(* Logix 5000 project; controller MECO9497 vendor 1 type 14 code 106 rev 21.11; software revision 21.00 *)

TASK MainTask (continuous, watchdog 500 ms) : MainProgram
TASK PID_LOOP (periodic, rate 250 ms, priority 5, watchdog 500 ms) : PID_MAIN
TASK PID_SLOW (periodic, rate 1000 ms, priority 10, watchdog 500 ms) : PID_SLOW

MODULES
   Local : vendor 1 type 14 code 106 (Compact 0, rev 21.11)
       : 1769-IQ16 (Compact 1, rev 1.1, Input RPI 20 ms)
       : 1769-IF8 (Compact 3, rev 1.1, Output RPI 80 ms)
       : vendor 1 type 10 code 40 (Compact 5, rev 2.1, Output RPI 80 ms)
       : 1769-OW16 (Compact 2, rev 1.1, Output RPI 20 ms)
       : 1769-IF8 (Compact 4, rev 1.1, Output RPI 80 ms)
END_MODULES

VAR_GLOBAL   (* controller tags *)
   AAH_200 : BOOL := 1;
   AAH_200_ACK : BOOL;
   AAH_200_AUX : BOOL := 1;
   AAH_200_DELAY : TIMER := (PRE := 1000);
   AAH_200_DI : ALIAS FOR Local:1:I.Data.5;
   AAH_200_SP : REAL := 0.6;
   AAH_200_SP_H : BOOL;
   AAH_200_SP_N : BOOL;
   AAH_200_SP_O : REAL := 0.6;
   ACKNOWLEDGE : BOOL;
   ALARM_ACK_OIT : BOOL;
   ALARM_HORN_DO : ALIAS FOR Local:2:O.Data.10;
   ALARM_RESET_OIT : BOOL;
   ALARM_SCREEN_DISPLAY_BIT : BOOL;
   ALARM_SCREEN_LATCH_BIT : BOOL;
   ALERT_ALARM_SU_DELAY : TIMER := (PRE := 300000);
   ALERT_ALARM_SU_DELAY_H : BOOL;
   ALERT_ALARM_SU_DELAY_N : BOOL;
   ALERT_ALARM_SU_DELAY_O : DINT := 300;
   AT_200_AI : ALIAS FOR Local:4:I.Ch0Data;
   AT_200_EU : REAL;
   AUDIBLE_SUMMARY : BOOL;
   COMP_AMP_ALRM_DELAY_TMR : TIMER := (PRE := 20000);
   COMP_BUMP_OIT : BOOL;
   COMP_BUMP_SU_DELAY : TIMER := (PRE := 20);
   COMPRESSOR_FAULT_DELAY : TIMER := (PRE := 3000);
   COMPRESSOR_MOTOR_FLT_STARTUP_DELAY : TIMER := (PRE := 6000);
   COMPRESSOR_MOTOR_START_DELAY : TIMER := (PRE := 5000);
   COMPRESSOR_MOTOR_START_DO : ALIAS FOR Local:2:O.Data.0;
   COMPRESSOR_START_CMD : BOOL;
   CR_4 : ALIAS FOR Local:2:O.Data.9;
   CR_6 : ALIAS FOR Local:2:O.Data.2;
   CURRENT_SCREEN : DINT := 7;
   D_V_ALERT_ALARM : BOOL;
   D_V_CRITICAL_ALARM : BOOL;
   D_V_OP_SWITCH_AUTO : BOOL := 1;
   D_V_OP_SWITCH_MAN : BOOL;
   D_V_OP_SWITCH_OFF : BOOL;
   D_V_REMOTE_START : BOOL;
   D_V_REMOTE_START_MAP : BOOL;
   D_V_UNIT_RUNNIING : BOOL;
   DELTA_V_FP : REAL[30] := ([2] := 0.006103888, [4] := 0.25801086, [5] := 100.0, [6] := 60.074467, [8] := 39.310135, [9] := 1.5030825, [11] := 40.0, [12] := 102.87493, [13] := 102.08753); {produced}
   DELTA_V_READ : INT[10] := ([0] := 2, [2] := 1344, [3] := 16383, [5] := 1); {produced}
   DELTA_V_WRITE : INT[10] := ([0] := 1); {produced}
   DIST_COND_ALRM_STARTUP_TIME_H : BOOL;
   DIST_COND_ALRM_STARTUP_TIME_N : BOOL;
   DIST_COND_ALRM_STARTUP_TIME_O : REAL := 300.0;
   DIST_COND_ALRM_STARTUP_TMR : TIMER := (PRE := 300000);
   DIST_MOTOR_BUMP_OIT : BOOL;
   DIST_PUMP_START_SP : REAL := 75.0;
   DIST_PUMP_START_SP_H : BOOL;
   DIST_PUMP_START_SP_N : BOOL;
   DIST_PUMP_START_SP_OIT : REAL := 80.0;
   DIST_PUMP_STOP_SP : REAL := 10.0;
   DIST_PUMP_STOP_SP_H : BOOL;
   DIST_PUMP_STOP_SP_N : BOOL;
   DIST_PUMP_STOP_SP_OIT : DINT := 20;
   DIST_TO_STORAGE_TIME_SP_H : BOOL;
   DIST_TO_STORAGE_TIME_SP_N : BOOL;
   DIST_TO_STORAGE_TIME_SP_OIT : DINT;
   DISTILATE_TO_STORAGE : BOOL;
   DISTILLATE_MOTOR_FAULT_DELAY : TIMER := (PRE := 3000);
   DISTILLATE_MOTOR_START_DO : ALIAS FOR Local:2:O.Data.1;
   DISTILLATE_PUMP_NORM_START : BOOL;
   DISTILLATE_PUMP_START_CMD : BOOL;
   DISTILLATE_PUMP_STDBY_START : BOOL;
   DSTLT_BOX_DRAIN_HOT_STANDBY : TIMER := (PRE := 600000, ACC := 600000, EN := 1, DN := 1);
   DSTLT_BOX_DRAIN_HOT_STANDBY_CLOSE : TIMER := (PRE := 1800000, ACC := 431720, EN := 1, TT := 1);
   DSTLT_BOX_DRAIN_NORM_DELAY : TIMER := (PRE := 5000);
   DSTLT_BOX_DRAIN_STANDBY : BOOL;
   DSTLT_BOX_DRAIN_STBY_DELAY_TIMER : TIMER := (PRE := 10000);
   DSTLT_PUMP_START_DELAY : TIMER := (PRE := 5000);
   DSTLT_PUMP_STBY_STOP_SP : REAL;
   DSTLT_PUMP_STBY_STRT_SP : REAL;
   DSTLT_STORAGE : BOOL;
   DSTLT_STORAGE_DELAY_TIMER : TIMER := (PRE := 60000);
   DSTLT_STORAGE_DELTA_V : BOOL;
   DSTLT_STORAGE_ENABLE_MAP : BOOL := 1;
   DSTLT_STORAGE_ENABLE_OIT : BOOL := 1;
   DSTLT_TEMP_ALRM_SU_DELAY : TIMER := (PRE := 300000);
   DSTLT_TEMP_ALRM_SU_DELAY_H : BOOL;
   DSTLT_TEMP_ALRM_SU_DELAY_N : BOOL;
   DSTLT_TEMP_ALRM_SU_DELAY_O : REAL := 300.0;
   DSTLT_TEMP_CNTRL_DELAY_TIMER : TIMER := (PRE := 90000);
   E_Stop : ALIAS FOR Local:1:I.Data.0;
   E_Stop_ACK : BOOL;
   E_Stop_AUX : BOOL := 1;
   E_Stop_DI_MAP : BOOL;
   ENGINEER : BOOL;
   EVAP_PRESS_CV_LIMIT : BOOL;
   EVAP_PRESS_CV_PERMISSIVE : REAL := 10.0;
   EVAP_PRESS_RAMP_ONE_SHOT : BOOL;
   EVAP_PRESS_RAMP_TIMER : TIMER := (PRE := 60000);
   EVAP_PRESSURE_CV_PERM : BOOL := 1;
   EVAP_PRESSURE_PERM : BOOL := 1;
   EVAP_PRESSURE_PERM_TIME_H : BOOL;
   EVAP_PRESSURE_PERM_TIME_N : BOOL;
   EVAP_PRESSURE_PERM_TIME_O : REAL := 180.0;
   EVAP_PRESSURE_PERM_TIMER : TIMER := (PRE := 180000, ACC := 180000, EN := 1, DN := 1);
   EVAP_RAMP_COMPLETE : BOOL;
   EVAP_RAMP_ENABLE_DELAY_TIMER : TIMER := (PRE := 180000);
   EXCESS_DIST_TIME_SP_H : BOOL;
   EXCESS_DIST_TIME_SP_N : BOOL;
   EXCESS_DIST_TIME_SP_OIT : REAL := 10.0;
   EXCESS_DIST_TO_DRAIN_ACK : BOOL;
   EXCESS_DIST_TO_DRAIN_AUX : BOOL := 1;
   EXCESS_DSTLT_DELAY_TIMER : TIMER := (PRE := 1000);
   EXCESS_DSTLT_DRAIN : BOOL := 1;
   EXCESS_DSTLT_DRAIN_TIMER : TIMER := (PRE := 600000);
   EXCESS_DSTLT_REMAIN : DINT := 10;
   FC_300_AM_OIT : BOOL;
   FC_300_OS_OFF : BOOL := 1;
   FC_300_OS_ON : BOOL;
   FC_300_SP : DINT := 58;
   FC_300_SP_H : BOOL;
   FC_300_SP_N : BOOL;
   FC_300_SP_O : DINT := 58;
   FC_300_SP_OUT : DINT;
   FEED_LVL_CV_LIMIT : BOOL := 1;
   FEED_LVL_CV_LIMIT_SHUTDOWN : BOOL := 1;
   FEED_LVL_CV_LIMIT_SHUTDOWN_DELAY : TIMER := (PRE := 30000);
   FEED_LVL_CV_LIMIT_SHUTDOWN_LATCH : BOOL;
   FEED_LVL_ONE_SHOT : BOOL;
   FEED_TEM_SD_LATCH : BOOL;
   FEED_TEM_SD_TIMER : TIMER := (PRE := 30000);
   FEED_TEMP_SD_ONS : BOOL := 1;
   FEED_TEMP_STEP_DELAY : TIMER := (PRE := 10000);
   FT_200_AI : ALIAS FOR Local:3:I.Ch2Data;
   FT_200_EU : REAL;
   HEARTBEAT : BOOL := 1;
   HEARTBEAT_AUX : BOOL;
   HEARTBEAT_OUT : BOOL := 1;
   HEARTBEAT_RESET_OIT : BOOL;
   HOT_STANDBY : BOOL := 1;
   HOURMETER_DO : ALIAS FOR Local:2:O.Data.4;
   IAL_100 : BOOL;
   IAL_100_ACK : BOOL;
   IAL_100_AUX : BOOL := 1;
   IAL_100_CTR : COUNTER := (PRE := 3);
   IAL_100_DELAY : TIMER := (PRE := 5000);
   IAL_100_SP : REAL := 30.0;
   IAL_100_SP_H : BOOL;
   IAL_100_SP_N : BOOL;
   IAL_100_SP_OIT : REAL := 30.0;
   INITIAL_SCAN_BIT : BOOL;
   INITIAL_SCAN_SYS_RESET : BOOL;
   INITIAL_SCAN_SYS_RESET_TMR : TIMER := (PRE := 30000);
   INITIAL_START_STEAM_LIMIT_TMR : TIMER := (PRE := 300000, ACC := 300000, EN := 1, DN := 1);
   IY_100_AI : ALIAS FOR Local:4:I.Ch2Data;
   IY_100_EU : REAL;
   LAAH_100 : BOOL := 1;
   LAAH_100_ACK : BOOL;
   LAAH_100_ALERT_H : BOOL;
   LAAH_100_ALERT_N : BOOL;
   LAAH_100_ALERT_O : DINT := 80;
   LAAH_100_AUX : BOOL := 1;
   LAAH_100_DELAY : TIMER := (PRE := 5000);
   LAAH_100_SP : DINT := 80;
   LAAL_100 : BOOL := 1;
   LAAL_100_ACK : BOOL;
   LAAL_100_ALERT_H : BOOL;
   LAAL_100_ALERT_N : BOOL;
   LAAL_100_ALERT_O : DINT := 20;
   LAAL_100_AUX : BOOL := 1;
   LAAL_100_DELAY : TIMER := (PRE := 1000);
   LAAL_100_SP : DINT := 20;
   LAH_100 : BOOL := 1;
   LAH_100_ACK : BOOL;
   LAH_100_AUX : BOOL := 1;
   LAH_100_DELAY : TIMER := (PRE := 5000);
   LAH_100_SP : REAL := 80.0;
   LAH_100_SP_H : BOOL;
   LAH_100_SP_N : BOOL;
   LAH_100_SP_OIT : REAL := 80.0;
   LAL_100 : BOOL := 1;
   LAL_100_ACK : BOOL;
   LAL_100_AUX : BOOL := 1;
   LAL_100_DELAY : TIMER := (PRE := 1000);
   LAL_100_SP : REAL := 20.0;
   LAL_100_SP_H : BOOL;
   LAL_100_SP_N : BOOL;
   LAL_100_SP_OIT : REAL := 20.0;
   LATCH : BOOL := 1;
   LB_OIL_LOW_PRESS_ALRM_DELAY : TIMER := (PRE := 20000);
   LCV_100_AO : ALIAS FOR Local:5:O.Ch2Data;
   LCV_100_IND : DINT;
   LCV_100_INTERLOCK : BOOL := 1;
   LCV_200_AO : ALIAS FOR Local:5:O.Ch3Data;
   LCV_200_IND : DINT := 3;
   LIC_100 : PID := (CTL := -2139061120, EN := 1, PE := 1, INI := 1, DVNA := 1, PVHA := 1, SP := 9829.8, KP := 4.0, KI := 1.6, KD := 0.01, BIAS := -181.60863, MAXS := 16383.0, SO := 0.25801086, MAXO := 40.0, UPD := 0.25, PV := 9845.0, ERR := -15.200195, OUT := 0.25801086, MAXI := 16383.0, MAXCV := 16383.0, MAXTIE := 16383.0, DATA[0] := 182.52715, DATA[1] := -961.19507, DATA[2] := 9845.0, DATA[3] := -15.200195, DATA[4] := 9829.8, DATA[5] := 0.006103888, DATA[6] := 1.0, DATA[7] := 6.3999996, DATA[8] := 4.0, DATA[9] := 1.6, DATA[10] := 0.01, DATA[11] := 4.0, DATA[12] := 0.041666668, DATA[13] := 2.3999999, DATA[15] := 163.83, DATA[16] := 0.006103888);
   LIC_1000_CV1 : REAL := 20.0;
   LIC_100_A_M_OIT : BOOL;
   LIC_100_CV2 : REAL := 40.0;
   LIC_100_CV_H : BOOL;
   LIC_100_CV_N : BOOL;
   LIC_100_CV_OIT : REAL := 0.25801086;
   LIC_100_FINAL_SP : REAL := 9829.8;
   LIC_100_FINAL_SP_EU : REAL := 60.0;
   LIC_100_GAIN_H : BOOL;
   LIC_100_GAIN_N : BOOL;
   LIC_100_GAIN_OIT : REAL := 4.0;
   LIC_100_RATE_H : BOOL;
   LIC_100_RATE_N : BOOL;
   LIC_100_RATE_OIT : REAL := 0.01;
   LIC_100_RESET_H : BOOL;
   LIC_100_RESET_N : BOOL;
   LIC_100_RESET_OIT : REAL := 1.6;
   LIC_100_SP_CONV : REAL := 163.83;
   LIC_100_SP_EU : REAL := 60.0;
   LIC_100_SP_H : BOOL;
   LIC_100_SP_N : BOOL;
   LIC_100_SP_OIT : REAL := 60.0;
   LIC_100_STBY_SP : REAL := 9829.8;
   LIC_100_STBY_SP_EU : REAL := 60.0;
   LIC_100_STBY_SP_H : BOOL;
   LIC_100_STBY_SP_N : BOOL;
   LIC_100_STBY_SP_OIT : REAL := 60.0;
   LIC_200 : PID := (CTL := -2038397696, EN := 1, SWM := 1, CA := 1, PE := 1, INI := 1, DVNA := 1, PVLA := 1, SP := 9829.8, KP := 2.0, KI := 1.1, KD := 0.01, BIAS := 151.65573, MAXS := 16383.0, SO := 100.0, MAXO := 100.0, UPD := 0.25, PV := -98.0, ERR := -9927.8, OUT := 100.0, MAXI := 16383.0, MAXCV := 16383.0, MAXTIE := 16383.0, DATA[0] := 69.54062, DATA[1] := -9.570896, DATA[2] := -98.0, DATA[3] := -9927.8, DATA[4] := 9829.8, DATA[5] := 0.006103888, DATA[6] := 1.0, DATA[7] := 5.2, DATA[8] := 2.0, DATA[9] := 1.1, DATA[10] := 0.01, DATA[11] := 2.0, DATA[12] := 0.030303031, DATA[13] := 1.1999999, DATA[15] := 163.83, DATA[16] := 0.006103888);
   LIC_200_A_M_OIT : BOOL;
   LIC_200_CV_H : BOOL;
   LIC_200_CV_N : BOOL;
   LIC_200_CV_OIT : REAL := 100.0;
   LIC_200_GAIN_H : BOOL;
   LIC_200_GAIN_N : BOOL;
   LIC_200_GAIN_OIT : REAL := 2.0;
   LIC_200_RATE_H : BOOL;
   LIC_200_RATE_N : BOOL;
   LIC_200_RATE_OIT : REAL := 0.01;
   LIC_200_RESET_H : BOOL;
   LIC_200_RESET_N : BOOL;
   LIC_200_RESET_OIT : REAL := 1.1;
   LIC_200_SP_CONV : REAL := 163.83;
   LIC_200_SP_EU : REAL := 60.0;
   LIC_200_SP_H : BOOL;
   LIC_200_SP_N : BOOL;
   LIC_200_SP_OIT : REAL := 60.0;
   LT_100_AI : ALIAS FOR Local:3:I.Ch3Data;
   LT_100_EU : REAL := 60.092777;
   LT_100_EU_SPAN : REAL := 100.0;
   LT_100_EU_ZERO : REAL;
   LT_200_AI : ALIAS FOR Local:3:I.Ch4Data;
   LT_200_EU : REAL;
   LT_200_EU_SPAN : REAL := 100.0;
   LT_200_EU_ZERO : REAL;
   LUBE_OIL_PUMP_FAULT_DELAY : TIMER := (PRE := 3000);
   LUBE_OIL_PUMP_START_CMD : BOOL;
   LUBE_OIL_SHUTDWN_TIMER : TIMER := (PRE := 45000, ACC := 45000, EN := 1, DN := 1);
   M1_DI : ALIAS FOR Local:1:I.Data.1;
   M1_DI_MAP : BOOL;
   M1_FAULT_ACK : BOOL;
   M1_FAULT_AUX : BOOL := 1;
   M2_DI : ALIAS FOR Local:1:I.Data.2;
   M2_DI_MAP : BOOL;
   M2_FAULT_ACK : BOOL;
   M2_FAULT_AUX : BOOL := 1;
   M4_DI : ALIAS FOR Local:1:I.Data.4;
   M4_DI_MAP : BOOL;
   M4_FAULT_ACK : BOOL;
   M4_FAULT_AUX : BOOL := 1;
   MAINTENANCE : BOOL;
   MCB : BOOL;
   MSG_AAH_200 : BOOL;
   MSG_E_STOP : BOOL;
   MSG_EXCESS_DIST_TO_DRAIN : BOOL;
   MSG_IAL_100 : BOOL;
   MSG_LAH_100 : BOOL;
   MSG_LAL_100 : BOOL;
   MSG_M1_FLT : BOOL;
   MSG_M2_FLT : BOOL;
   MSG_M4_FLT : BOOL;
   MSG_PAH_103 : BOOL;
   MSG_PAL_103 : BOOL;
   MSG_PAL_700 : BOOL;
   MSG_TAH_700 : BOOL;
   MSG_TAL_200 : BOOL;
   MSS_ALERT : BOOL;
   MSS_AUTO_SHUTDOWN_LATCH : BOOL;
   MSS_SHUTDOWN : BOOL := 1;
   MSS_START_PERM : BOOL := 1;
   no : BOOL;
   OFF : BOOL;
   OIL_MOTOR_START_DO : ALIAS FOR Local:2:O.Data.11;
   OIT_SCREEN_CONTROL : DINT;
   OIT_SECURITY_LEVEL : DINT;
   OP_SWTCH_AUTO_DI : ALIAS FOR Local:1:I.Data.14;
   OP_SWTCH_AUTO_DI_MAP : BOOL := 1;
   OP_SWTCH_MANUAL_DI : ALIAS FOR Local:1:I.Data.13;
   OP_SWTCH_MANUAL_DI_MAP : BOOL;
   OPERATOR : BOOL;
   PAAH_103 : BOOL := 1;
   PAAH_103_ACK : BOOL;
   PAAH_103_ALERT_H : BOOL;
   PAAH_103_ALERT_N : BOOL;
   PAAH_103_ALERT_O : REAL := 3.0;
   PAAH_103_AUX : BOOL := 1;
   PAAH_103_DELAY : TIMER := (PRE := 1000);
   PAAH_103_SP : REAL := 3.0;
   PAAL_103 : BOOL := 1;
   PAAL_103_ACK : BOOL;
   PAAL_103_ALERT_H : BOOL;
   PAAL_103_ALERT_N : BOOL;
   PAAL_103_ALERT_O : REAL := 0.25;
   PAAL_103_AUX : BOOL := 1;
   PAAL_103_DELAY : TIMER := (PRE := 1000);
   PAAL_103_SP : REAL := 0.25;
   PAH_103 : BOOL := 1;
   PAH_103_ACK : BOOL;
   PAH_103_AUX : BOOL := 1;
   PAH_103_DELAY : TIMER := (PRE := 1000);
   PAH_103_SP : REAL := 3.0;
   PAH_103_SP_H : BOOL;
   PAH_103_SP_N : BOOL;
   PAH_103_SP_OIT : REAL := 3.0;
   PAL_103 : BOOL := 1;
   PAL_103_ACK : BOOL;
   PAL_103_AUX : BOOL := 1;
   PAL_103_DELAY : TIMER := (PRE := 1000);
   PAL_103_SP : REAL := 0.19;
   PAL_103_SP_H : BOOL;
   PAL_103_SP_N : BOOL;
   PAL_103_SP_OIT : REAL := 0.19;
   PAL_700 : BOOL;
   PAL_700_ACK : BOOL;
   PAL_700_ALRM_DELAY : TIMER := (PRE := 1000);
   PAL_700_AUX : BOOL := 1;
   PCV_103_AO : ALIAS FOR Local:5:O.Ch0Data;
   PCV_103_IND : DINT := 3;
   PCV_103_INTERLOCK : BOOL := 1;
   PERM_TIME_REMAINING : REAL;
   PIC_103 : PID := (CTL := -2139061120, EN := 1, PE := 1, INI := 1, DVNA := 1, PVHA := 1, SP := 4914.9004, KP := 3.5, KI := 1.0, KD := 0.01, BIAS := -117.88922, MAXS := 16383.0, SO := 39.310135, MAXO := 100.0, UPD := 0.25, PV := 4920.0, ERR := -5.0996094, OUT := 39.310135, MAXI := 16383.0, MAXCV := 16383.0, MAXTIE := 16383.0, DATA[0] := 157.11327, DATA[1] := -480.6931, DATA[2] := 4920.0, DATA[3] := -5.0996094, DATA[4] := 4914.9004, DATA[5] := 0.006103888, DATA[6] := 1.0, DATA[7] := 6.1, DATA[8] := 3.5, DATA[9] := 1.0, DATA[10] := 0.01, DATA[11] := 3.5, DATA[12] := 0.058333334, DATA[13] := 2.1, DATA[15] := 163.83, DATA[16] := 0.006103888);
   PIC_103_A_M_OIT : BOOL;
   PIC_103_CV_H : BOOL;
   PIC_103_CV_N : BOOL;
   PIC_103_CV_OIT : REAL := 38.848907;
   PIC_103_FINAL_SP : REAL := 1.0;
   PIC_103_GAIN_H : BOOL;
   PIC_103_GAIN_N : BOOL;
   PIC_103_GAIN_OIT : REAL := 3.5;
   PIC_103_RATE_H : BOOL;
   PIC_103_RATE_N : BOOL;
   PIC_103_RATE_OIT : REAL := 0.01;
   PIC_103_RESET_H : BOOL;
   PIC_103_RESET_N : BOOL;
   PIC_103_RESET_OIT : REAL := 1.0;
   PIC_103_SP_CONV : REAL := 3276.6;
   PIC_103_SP_EU : REAL := 1.5000001;
   PIC_103_SP_H : BOOL;
   PIC_103_SP_N : BOOL;
   PIC_103_SP_OIT : REAL := 1.0;
   PIC_103_STBY_SP : REAL := 4914.9004;
   PIC_103_STBY_SP_EU : REAL := 1.5000001;
   PIC_103_STBY_SP_H : BOOL;
   PIC_103_STBY_SP_N : BOOL;
   PIC_103_STBY_SP_OIT : REAL := 1.5;
   PSL_700_DI : ALIAS FOR Local:1:I.Data.7;
   PT_103_AI : ALIAS FOR Local:3:I.Ch0Data;
   PT_103_EU : REAL := 1.5015565;
   PT_103_EU_SPAN : REAL := 5.0;
   PT_103_EU_ZERO : REAL;
   PT_103_HIGH : REAL := 2.1;
   RESET : BOOL;
   RESET_CONDUCTIVITY_HIGH_OIT : BOOL;
   RESET_DIST_LOW_TEMP_OIT : BOOL;
   SECURITY_ENABLED : BOOL;
   SUPERVISOR : BOOL;
   SV_200 : ALIAS FOR Local:2:O.Data.5;
   SV_200_201_DO : ALIAS FOR Local:2:O.Data.6;
   SV_200_201_IND : BOOL;
   SV_200_CTL : BOOL;
   SV_200_IND : BOOL;
   SV_202_DO : ALIAS FOR Local:2:O.Data.5;
   SV_300_DO : ALIAS FOR Local:2:O.Data.3;
   SV_300_IND : BOOL;
   SV_500_DO : ALIAS FOR Local:2:O.Data.8;
   SV_500_IND : BOOL;
   TAH_700 : BOOL := 1;
   TAH_700_ACK : BOOL;
   TAH_700_ALRM_DELAY : TIMER := (PRE := 3000);
   TAH_700_AUX : BOOL := 1;
   TAL_200 : BOOL := 1;
   TAL_200_ACK : BOOL;
   TAL_200_AUX : BOOL := 1;
   TAL_200_DELAY : TIMER := (PRE := 10000);
   TAL_200_SP : REAL := 76.0;
   TAL_200_SP_H : BOOL;
   TAL_200_SP_N : BOOL;
   TAL_200_SP_OIT : REAL := 76.0;
   TCV_102_AO : ALIAS FOR Local:5:O.Ch4Data;
   TCV_102_IND : DINT;
   TCV_200_AO : ALIAS FOR Local:5:O.Ch1Data;
   TCV_200_IND : DINT := 3;
   test : BOOL;
   TIC_102 : PID := (CTL := -2071952256, EN := 1, SWM := 1, PE := 1, INI := 1, DVNA := 1, PVHA := 1, SP := 11031.22, KP := 2.5, KI := 1.0, KD := 0.02, BIAS := -106.50499, MAXS := 16383.0, MAXO := 100.0, UPD := 1.0, PV := 11236.0, ERR := -204.78027, MAXI := 16383.0, MAXCV := 16383.0, MAXTIE := 16383.0, DATA[0] := 109.65634, DATA[1] := -1097.3062, DATA[2] := 11236.0, DATA[3] := -204.78027, DATA[4] := 11031.22, DATA[5] := 0.006103888, DATA[6] := 1.0, DATA[7] := 19.0, DATA[8] := 2.5, DATA[9] := 1.0, DATA[10] := 0.02, DATA[11] := 2.5, DATA[12] := 0.041666668, DATA[13] := 2.9999998, DATA[15] := 163.83, DATA[16] := 0.006103888);
   TIC_102_A_M_OIT : BOOL;
   TIC_102_CV_H : BOOL;
   TIC_102_CV_MIN_LIMIT : BOOL;
   TIC_102_CV_N : BOOL;
   TIC_102_CV_OIT : REAL;
   TIC_102_CV_SU_H : BOOL;
   TIC_102_CV_SU_N : BOOL;
   TIC_102_CV_SU_O : DINT := 40;
   TIC_102_CV_SU_REM : DINT := 120;
   TIC_102_CV_SU_TIMER : TIMER := (PRE := 120000);
   TIC_102_GAIN_H : BOOL;
   TIC_102_GAIN_N : BOOL;
   TIC_102_GAIN_OIT : REAL := 2.5;
   TIC_102_MINCV1 : REAL := 20.0;
   TIC_102_MINCV2 : REAL := 40.0;
   TIC_102_MINCV3 : REAL := 60.0;
   TIC_102_RATE_H : BOOL;
   TIC_102_RATE_N : BOOL;
   TIC_102_RATE_OIT : REAL := 0.02;
   TIC_102_RESET_H : BOOL;
   TIC_102_RESET_N : BOOL;
   TIC_102_RESET_OIT : REAL := 1.0;
   TIC_102_SP_CONV : REAL := 109.22;
   TIC_102_SP_EU : REAL := 101.0;
   TIC_102_SP_H : BOOL;
   TIC_102_SP_N : BOOL;
   TIC_102_SP_OIT : REAL := 101.0;
   TIC_102_START_CV_TIMER_SP_H : BOOL;
   TIC_102_START_CV_TIMER_SP_N : BOOL;
   TIC_102_START_CV_TIMER_SP_O : REAL := 120.0;
   TIC_200 : PID := (CTL := -2071952256, EN := 1, SWM := 1, PE := 1, INI := 1, DVNA := 1, PVHA := 1, SP := 9065.26, KP := 4.5, KI := 1.0, KD := 0.02, BIAS := -92.58263, MAXS := 16383.0, SO := 40.0, MAXO := 100.0, UPD := 1.0, PV := 11142.0, ERR := -2076.7402, OUT := 40.0, MAXI := 16383.0, MAXCV := 16383.0, MAXTIE := 16383.0, DATA[0] := 189.52979, DATA[1] := -1088.248, DATA[2] := 11142.0, DATA[3] := -2076.7402, DATA[4] := 9065.26, DATA[5] := 0.006103888, DATA[6] := 1.0, DATA[7] := 21.4, DATA[8] := 4.5, DATA[9] := 1.0, DATA[10] := 0.02, DATA[11] := 4.5, DATA[12] := 0.075, DATA[13] := 5.3999996, DATA[15] := 163.83, DATA[16] := 0.006103888);
   TIC_200_A_M_OIT : BOOL;
   TIC_200_CV_H : BOOL;
   TIC_200_CV_N : BOOL;
   TIC_200_CV_OIT : REAL := 40.0;
   TIC_200_GAIN_H : BOOL;
   TIC_200_GAIN_N : BOOL;
   TIC_200_GAIN_OIT : REAL := 4.5;
   TIC_200_PER_OPEN : REAL := 60.0;
   TIC_200_RATE_H : BOOL;
   TIC_200_RATE_N : BOOL;
   TIC_200_RATE_OIT : REAL := 0.02;
   TIC_200_RESET_H : BOOL;
   TIC_200_RESET_N : BOOL;
   TIC_200_RESET_OIT : REAL := 1.0;
   TIC_200_SP_CONV : REAL := 109.22;
   TIC_200_SP_EU : REAL := 83.0;
   TIC_200_SP_H : BOOL;
   TIC_200_SP_N : BOOL;
   TIC_200_SP_OIT : REAL := 60.0;
   TIMER_BIT : TIMER := (PRE := 1000, ACC := 1000, EN := 1, DN := 1);
   TIMER_OUT : TIMER := (PRE := 5000, ACC := 366, EN := 1, TT := 1);
   TSH_700_DI : ALIAS FOR Local:1:I.Data.8;
   TT_102_AI : ALIAS FOR Local:3:I.Ch1Data;
   TT_102_EU : REAL := 102.85662;
   TT_102_EU_SPAN : REAL := 150.0;
   TT_102_EU_ZERO : REAL;
   TT_200_AI : ALIAS FOR Local:4:I.Ch1Data;
   TT_200_EU : REAL := 101.99597;
   TT_200_EU_SPAN : REAL := 150.0;
   TT_200_EU_ZERO : REAL;
   UNIT_REMOTE_START_DI : ALIAS FOR Local:1:I.Data.12;
   UNIT_REMOTE_START_MAP : BOOL;
   UNIT_START_DI : ALIAS FOR Local:1:I.Data.10;
   UNIT_START_DI_MAP : BOOL;
   UNIT_STATUS : DINT := 1;
   UNIT_STOP_DI : ALIAS FOR Local:1:I.Data.11;
   UNIT_STOP_DI_MAP : BOOL := 1;
END_VAR

PROGRAM MainProgram   (* main routine MainRoutine *)
VAR
   AT_200_SCALE : SCALE := (In := -97.0, InRawMax := 16383.0, InEUMax := 3.0, Limiting := 1, MinAlarm := 1);
   COM_LOW_BIT : BOOL;
   FT_200_SCALE : SCALE := (In := 4.0, InRawMax := 16383.0, InEUMax := 50.0, Limiting := 1, Out := 0.012207776);
   IY_100_SCALE : SCALE := (In := 49.0, InRawMax := 16383.0, InEUMax := 100.0, Limiting := 1, Out := 0.2990905);
   LOSS_COM_DISPLAY : TIMER := (PRE := 10000, ACC := 601, EN := 1, TT := 1);
   LT_100_SCALE : SCALE := (In := 9838.0, InRawMax := 16383.0, InEUMax := 100.0, Limiting := 1, Out := 60.050053);
   LT_200_SCALE : SCALE := (In := -98.0, InRawMax := 16383.0, InEUMax := 100.0, Limiting := 1, MinAlarm := 1);
   PT_103_SCALE : SCALE := (In := 4929.0, InRawMax := 16383.0, InEUMax := 5.0, Limiting := 1, Out := 1.5043032);
   SCL_01 : SCALE;
   TT_102_SCALE : SCALE := (In := 11237.0, InRawMax := 16383.0, InEUMax := 150.0, Limiting := 1, Out := 102.88409);
   TT_200_SCALE : SCALE := (In := 11144.0, InRawMax := 16383.0, InEUMax := 150.0, Limiting := 1, Out := 102.03259);
END_VAR

ROUTINE ALARMS   (* ladder *)
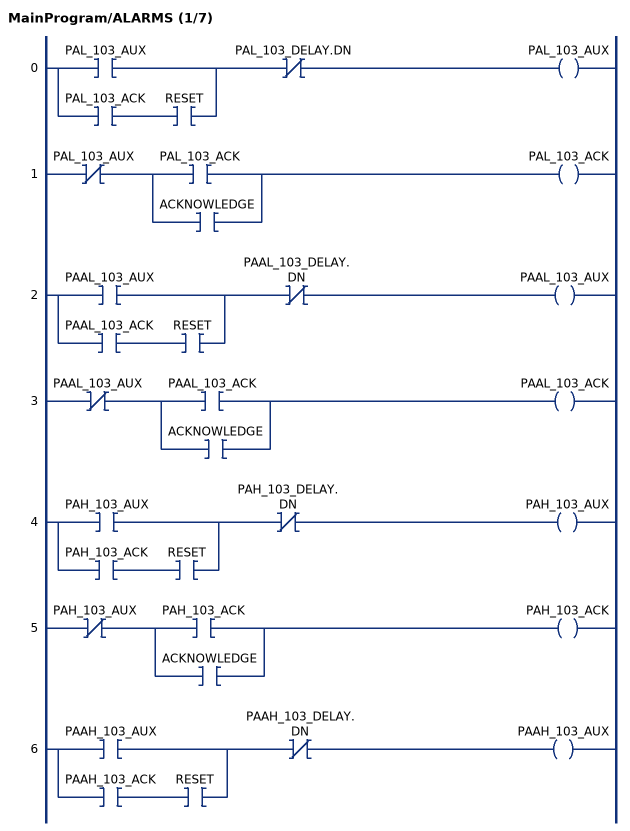
   0: [XIC(PAL_103_AUX) ,XIC(PAL_103_ACK) XIC(RESET) ]XIO(PAL_103_DELAY.DN)OTE(PAL_103_AUX);
   1: XIO(PAL_103_AUX)[XIC(PAL_103_ACK) ,XIC(ACKNOWLEDGE) ]OTE(PAL_103_ACK);
   2: [XIC(PAAL_103_AUX) ,XIC(PAAL_103_ACK) XIC(RESET) ]XIO(PAAL_103_DELAY.DN)OTE(PAAL_103_AUX);
   3: XIO(PAAL_103_AUX)[XIC(PAAL_103_ACK) ,XIC(ACKNOWLEDGE) ]OTE(PAAL_103_ACK);
   4: [XIC(PAH_103_AUX) ,XIC(PAH_103_ACK) XIC(RESET) ]XIO(PAH_103_DELAY.DN)OTE(PAH_103_AUX);
   5: XIO(PAH_103_AUX)[XIC(PAH_103_ACK) ,XIC(ACKNOWLEDGE) ]OTE(PAH_103_ACK);
   6: [XIC(PAAH_103_AUX) ,XIC(PAAH_103_ACK) XIC(RESET) ]XIO(PAAH_103_DELAY.DN)OTE(PAAH_103_AUX);
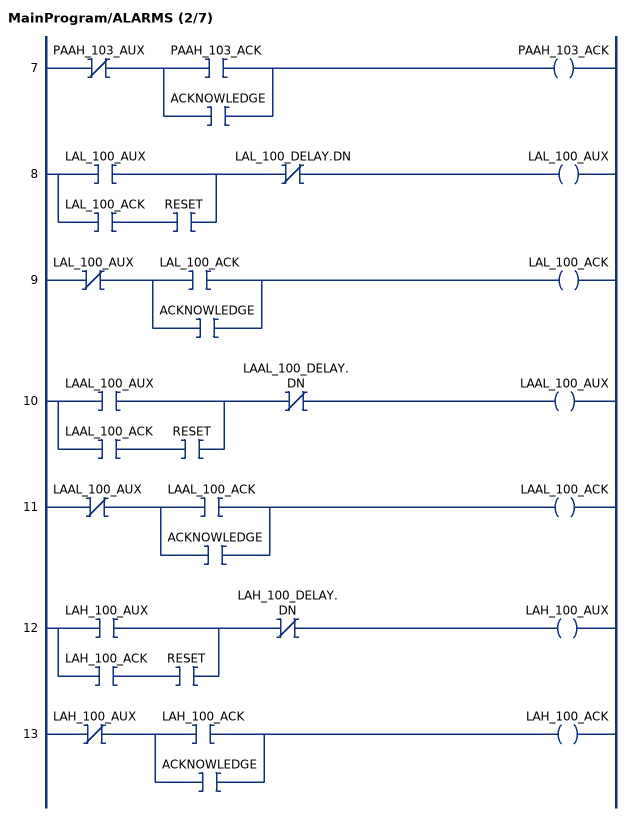
   7: XIO(PAAH_103_AUX)[XIC(PAAH_103_ACK) ,XIC(ACKNOWLEDGE) ]OTE(PAAH_103_ACK);
   8: [XIC(LAL_100_AUX) ,XIC(LAL_100_ACK) XIC(RESET) ]XIO(LAL_100_DELAY.DN)OTE(LAL_100_AUX);
   9: XIO(LAL_100_AUX)[XIC(LAL_100_ACK) ,XIC(ACKNOWLEDGE) ]OTE(LAL_100_ACK);
   10: [XIC(LAAL_100_AUX) ,XIC(LAAL_100_ACK) XIC(RESET) ]XIO(LAAL_100_DELAY.DN)OTE(LAAL_100_AUX);
   11: XIO(LAAL_100_AUX)[XIC(LAAL_100_ACK) ,XIC(ACKNOWLEDGE) ]OTE(LAAL_100_ACK);
   12: [XIC(LAH_100_AUX) ,XIC(LAH_100_ACK) XIC(RESET) ]XIO(LAH_100_DELAY.DN)OTE(LAH_100_AUX);
   13: XIO(LAH_100_AUX)[XIC(LAH_100_ACK) ,XIC(ACKNOWLEDGE) ]OTE(LAH_100_ACK);
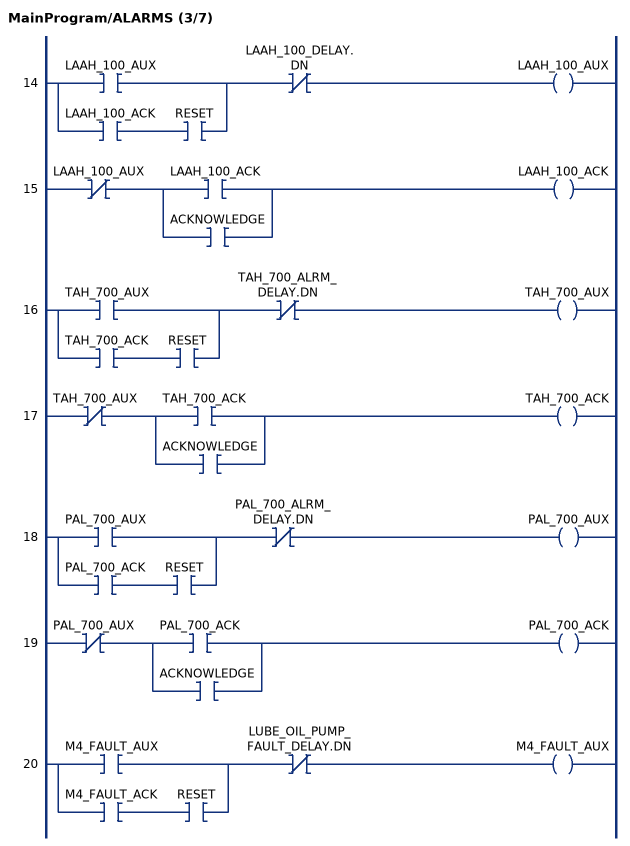
   14: [XIC(LAAH_100_AUX) ,XIC(LAAH_100_ACK) XIC(RESET) ]XIO(LAAH_100_DELAY.DN)OTE(LAAH_100_AUX);
   15: XIO(LAAH_100_AUX)[XIC(LAAH_100_ACK) ,XIC(ACKNOWLEDGE) ]OTE(LAAH_100_ACK);
   16: [XIC(TAH_700_AUX) ,XIC(TAH_700_ACK) XIC(RESET) ]XIO(TAH_700_ALRM_DELAY.DN)OTE(TAH_700_AUX);
   17: XIO(TAH_700_AUX)[XIC(TAH_700_ACK) ,XIC(ACKNOWLEDGE) ]OTE(TAH_700_ACK);
   18: [XIC(PAL_700_AUX) ,XIC(PAL_700_ACK) XIC(RESET) ]XIO(PAL_700_ALRM_DELAY.DN)OTE(PAL_700_AUX);
   19: XIO(PAL_700_AUX)[XIC(PAL_700_ACK) ,XIC(ACKNOWLEDGE) ]OTE(PAL_700_ACK);
   20: [XIC(M4_FAULT_AUX) ,XIC(M4_FAULT_ACK) XIC(RESET) ]XIO(LUBE_OIL_PUMP_FAULT_DELAY.DN)OTE(M4_FAULT_AUX);
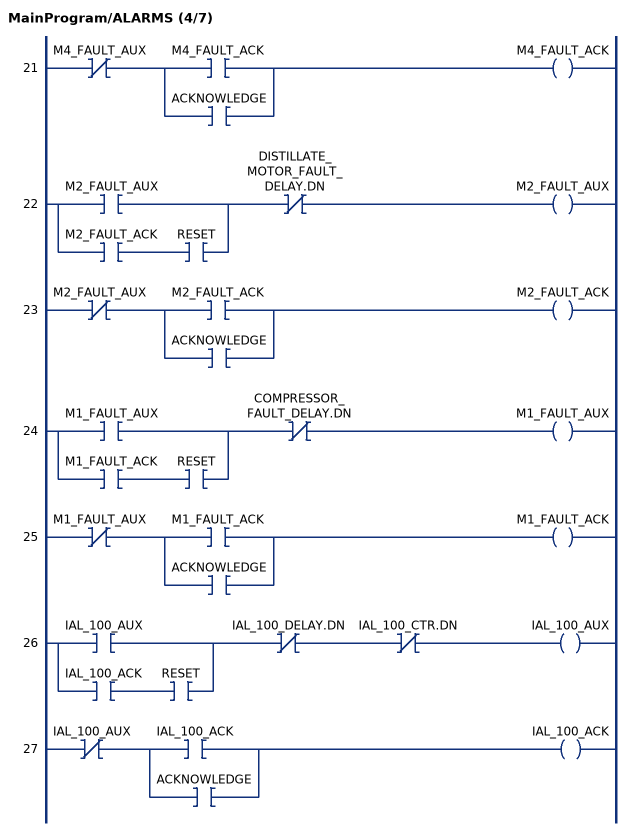
   21: XIO(M4_FAULT_AUX)[XIC(M4_FAULT_ACK) ,XIC(ACKNOWLEDGE) ]OTE(M4_FAULT_ACK);
   22: [XIC(M2_FAULT_AUX) ,XIC(M2_FAULT_ACK) XIC(RESET) ]XIO(DISTILLATE_MOTOR_FAULT_DELAY.DN)OTE(M2_FAULT_AUX);
   23: XIO(M2_FAULT_AUX)[XIC(M2_FAULT_ACK) ,XIC(ACKNOWLEDGE) ]OTE(M2_FAULT_ACK);
   24: [XIC(M1_FAULT_AUX) ,XIC(M1_FAULT_ACK) XIC(RESET) ]XIO(COMPRESSOR_FAULT_DELAY.DN)OTE(M1_FAULT_AUX);
   25: XIO(M1_FAULT_AUX)[XIC(M1_FAULT_ACK) ,XIC(ACKNOWLEDGE) ]OTE(M1_FAULT_ACK);
   26: [XIC(IAL_100_AUX) ,XIC(IAL_100_ACK) XIC(RESET) ]XIO(IAL_100_DELAY.DN)XIO(IAL_100_CTR.DN)OTE(IAL_100_AUX);
   27: XIO(IAL_100_AUX)[XIC(IAL_100_ACK) ,XIC(ACKNOWLEDGE) ]OTE(IAL_100_ACK);
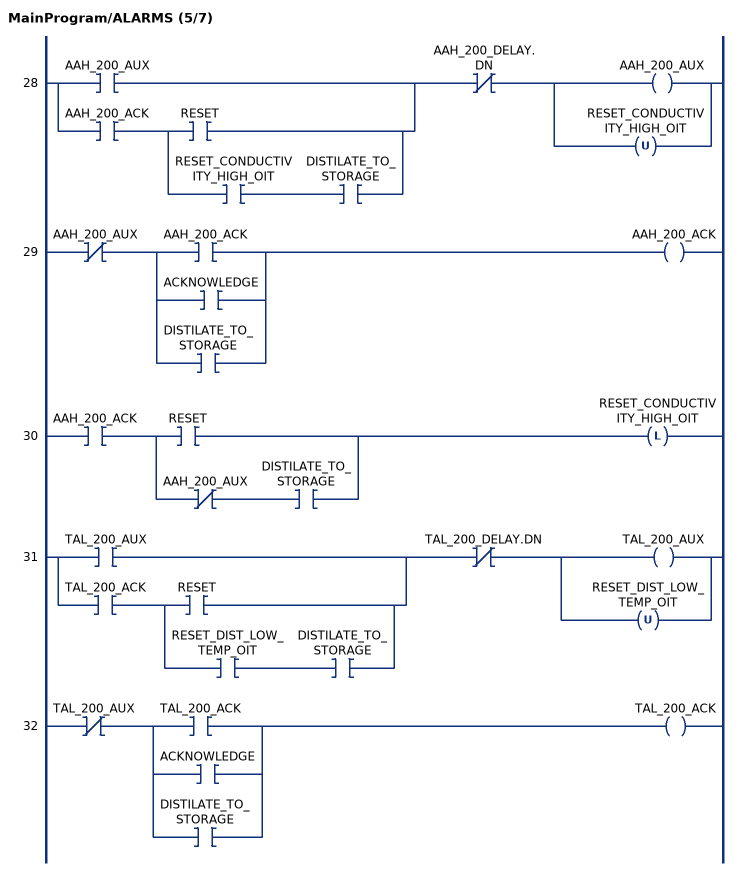
   28: [XIC(AAH_200_AUX) ,XIC(AAH_200_ACK) [XIC(RESET) ,XIC(RESET_CONDUCTIVITY_HIGH_OIT) XIC(DISTILATE_TO_STORAGE) ] ]XIO(AAH_200_DELAY.DN)[OTE(AAH_200_AUX) ,OTU(RESET_CONDUCTIVITY_HIGH_OIT) ];
   29: XIO(AAH_200_AUX)[XIC(AAH_200_ACK) ,XIC(ACKNOWLEDGE) ,XIC(DISTILATE_TO_STORAGE) ]OTE(AAH_200_ACK);
   30: XIC(AAH_200_ACK)[XIC(RESET) ,XIO(AAH_200_AUX) XIC(DISTILATE_TO_STORAGE) ]OTL(RESET_CONDUCTIVITY_HIGH_OIT);
   31: [XIC(TAL_200_AUX) ,XIC(TAL_200_ACK) [XIC(RESET) ,XIC(RESET_DIST_LOW_TEMP_OIT) XIC(DISTILATE_TO_STORAGE) ] ]XIO(TAL_200_DELAY.DN)[OTE(TAL_200_AUX) ,OTU(RESET_DIST_LOW_TEMP_OIT) ];
   32: XIO(TAL_200_AUX)[XIC(TAL_200_ACK) ,XIC(ACKNOWLEDGE) ,XIC(DISTILATE_TO_STORAGE) ]OTE(TAL_200_ACK);
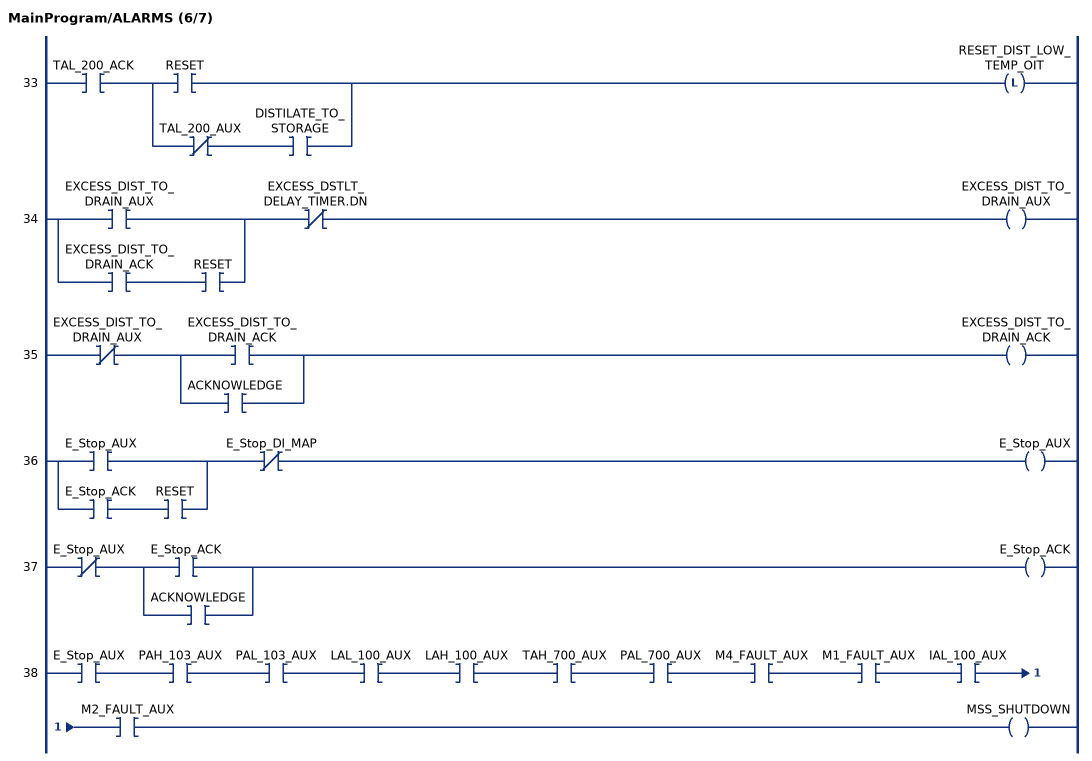
   33: XIC(TAL_200_ACK)[XIC(RESET) ,XIO(TAL_200_AUX) XIC(DISTILATE_TO_STORAGE) ]OTL(RESET_DIST_LOW_TEMP_OIT);
   34: [XIC(EXCESS_DIST_TO_DRAIN_AUX) ,XIC(EXCESS_DIST_TO_DRAIN_ACK) XIC(RESET) ]XIO(EXCESS_DSTLT_DELAY_TIMER.DN)OTE(EXCESS_DIST_TO_DRAIN_AUX);
   35: XIO(EXCESS_DIST_TO_DRAIN_AUX)[XIC(EXCESS_DIST_TO_DRAIN_ACK) ,XIC(ACKNOWLEDGE) ]OTE(EXCESS_DIST_TO_DRAIN_ACK);
   36: [XIC(E_Stop_AUX) ,XIC(E_Stop_ACK) XIC(RESET) ]XIO(E_Stop_DI_MAP)OTE(E_Stop_AUX);
   37: XIO(E_Stop_AUX)[XIC(E_Stop_ACK) ,XIC(ACKNOWLEDGE) ]OTE(E_Stop_ACK);
   38: XIC(E_Stop_AUX)XIC(PAH_103_AUX)XIC(PAL_103_AUX)XIC(LAL_100_AUX)XIC(LAH_100_AUX)XIC(TAH_700_AUX)XIC(PAL_700_AUX)XIC(M4_FAULT_AUX)XIC(M1_FAULT_AUX)XIC(IAL_100_AUX)XIC(M2_FAULT_AUX)OTE(MSS_SHUTDOWN);
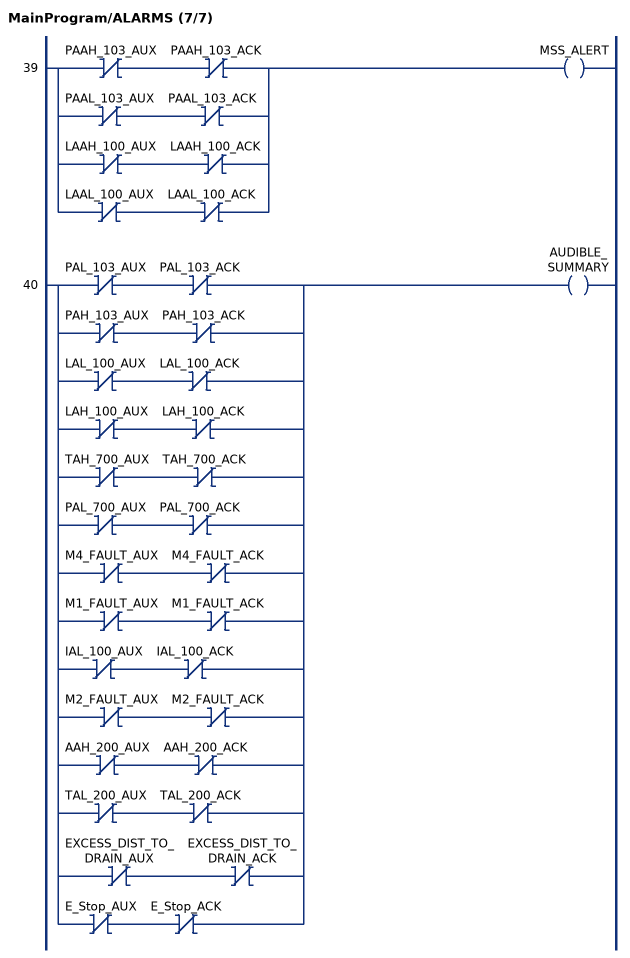
   39: [XIO(PAAH_103_AUX) XIO(PAAH_103_ACK) ,XIO(PAAL_103_AUX) XIO(PAAL_103_ACK) ,XIO(LAAH_100_AUX) XIO(LAAH_100_ACK) ,XIO(LAAL_100_AUX) XIO(LAAL_100_ACK) ]OTE(MSS_ALERT);
   40: [XIO(PAL_103_AUX) XIO(PAL_103_ACK) ,XIO(PAH_103_AUX) XIO(PAH_103_ACK) ,XIO(LAL_100_AUX) XIO(LAL_100_ACK) ,XIO(LAH_100_AUX) XIO(LAH_100_ACK) ,XIO(TAH_700_AUX) XIO(TAH_700_ACK) ,XIO(PAL_700_AUX) XIO(PAL_700_ACK) ,XIO(M4_FAULT_AUX) XIO(M4_FAULT_ACK) ,XIO(M1_FAULT_AUX) XIO(M1_FAULT_ACK) ,XIO(IAL_100_AUX) XIO(IAL_100_ACK) ,XIO(M2_FAULT_AUX) XIO(M2_FAULT_ACK) ,XIO(AAH_200_AUX) XIO(AAH_200_ACK) ,XIO(TAL_200_AUX) XIO(TAL_200_ACK) ,XIO(EXCESS_DIST_TO_DRAIN_AUX) XIO(EXCESS_DIST_TO_DRAIN_ACK) ,XIO(E_Stop_AUX) XIO(E_Stop_ACK) ]OTE(AUDIBLE_SUMMARY);
END_ROUTINE

ROUTINE DELTA_V   (* ladder *)
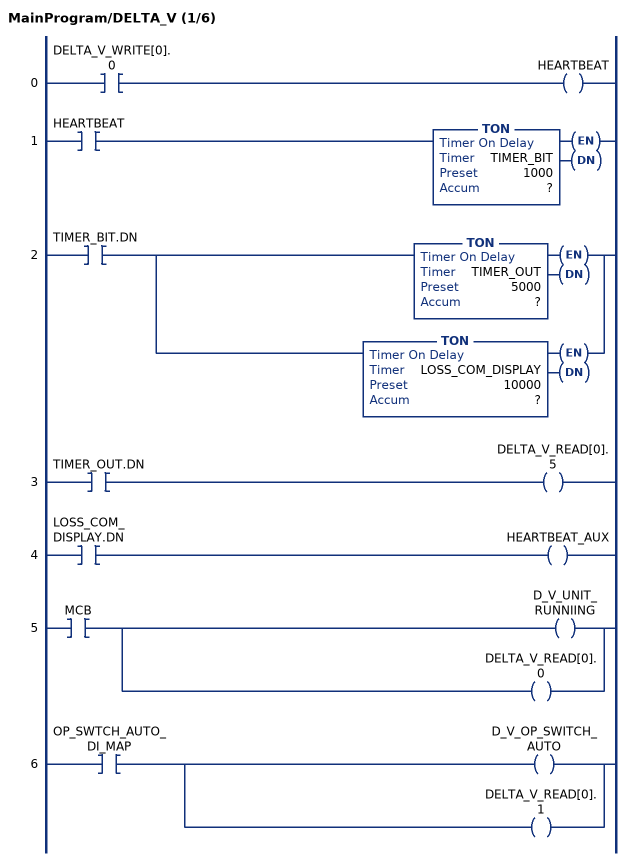
   0: XIC(DELTA_V_WRITE[0].0)OTE(HEARTBEAT);
   1: XIC(HEARTBEAT)TON(TIMER_BIT,?,?);
   2: XIC(TIMER_BIT.DN)[TON(TIMER_OUT,?,?) ,TON(LOSS_COM_DISPLAY,?,?) ];
   3: XIC(TIMER_OUT.DN)OTE(DELTA_V_READ[0].5);
   4: XIC(LOSS_COM_DISPLAY.DN)OTE(HEARTBEAT_AUX);
   5: XIC(MCB)[OTE(D_V_UNIT_RUNNIING) ,OTE(DELTA_V_READ[0].0) ];
   6: XIC(OP_SWTCH_AUTO_DI_MAP)[OTE(D_V_OP_SWITCH_AUTO) ,OTE(DELTA_V_READ[0].1) ];
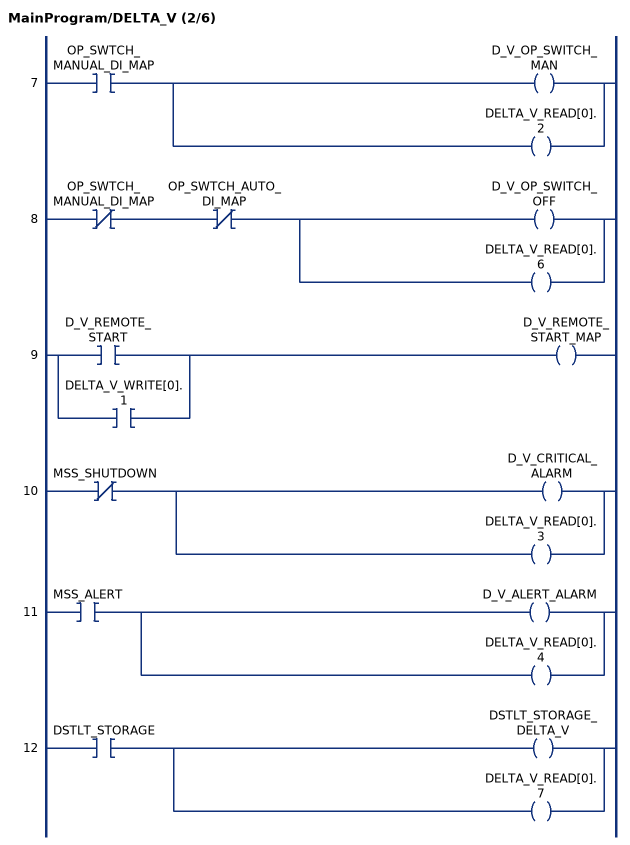
   7: XIC(OP_SWTCH_MANUAL_DI_MAP)[OTE(D_V_OP_SWITCH_MAN) ,OTE(DELTA_V_READ[0].2) ];
   8: XIO(OP_SWTCH_MANUAL_DI_MAP)XIO(OP_SWTCH_AUTO_DI_MAP)[OTE(D_V_OP_SWITCH_OFF) ,OTE(DELTA_V_READ[0].6) ];
   9: [XIC(D_V_REMOTE_START) ,XIC(DELTA_V_WRITE[0].1) ]OTE(D_V_REMOTE_START_MAP);
   10: XIO(MSS_SHUTDOWN)[OTE(D_V_CRITICAL_ALARM) ,OTE(DELTA_V_READ[0].3) ];
   11: XIC(MSS_ALERT)[OTE(D_V_ALERT_ALARM) ,OTE(DELTA_V_READ[0].4) ];
   12: XIC(DSTLT_STORAGE)[OTE(DSTLT_STORAGE_DELTA_V) ,OTE(DELTA_V_READ[0].7) ];
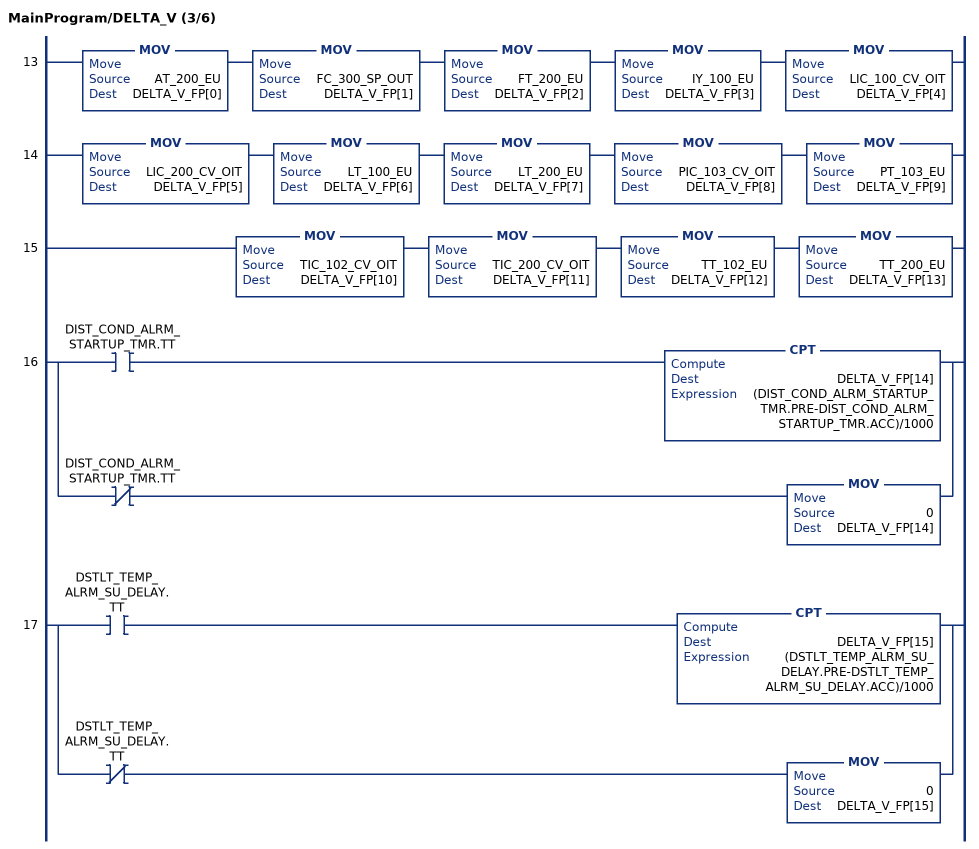
   13: MOV(AT_200_EU,DELTA_V_FP[0])MOV(FC_300_SP_OUT,DELTA_V_FP[1])MOV(FT_200_EU,DELTA_V_FP[2])MOV(IY_100_EU,DELTA_V_FP[3])MOV(LIC_100_CV_OIT,DELTA_V_FP[4]);
   14: MOV(LIC_200_CV_OIT,DELTA_V_FP[5])MOV(LT_100_EU,DELTA_V_FP[6])MOV(LT_200_EU,DELTA_V_FP[7])MOV(PIC_103_CV_OIT,DELTA_V_FP[8])MOV(PT_103_EU,DELTA_V_FP[9]);
   15: MOV(TIC_102_CV_OIT,DELTA_V_FP[10])MOV(TIC_200_CV_OIT,DELTA_V_FP[11])MOV(TT_102_EU,DELTA_V_FP[12])MOV(TT_200_EU,DELTA_V_FP[13]);
   16: [XIC(DIST_COND_ALRM_STARTUP_TMR.TT) CPT(DELTA_V_FP[14],(DIST_COND_ALRM_STARTUP_TMR.PRE-DIST_COND_ALRM_STARTUP_TMR.ACC)/1000) ,XIO(DIST_COND_ALRM_STARTUP_TMR.TT) MOV(0,DELTA_V_FP[14]) ];
   17: [XIC(DSTLT_TEMP_ALRM_SU_DELAY.TT) CPT(DELTA_V_FP[15],(DSTLT_TEMP_ALRM_SU_DELAY.PRE-DSTLT_TEMP_ALRM_SU_DELAY.ACC)/1000) ,XIO(DSTLT_TEMP_ALRM_SU_DELAY.TT) MOV(0,DELTA_V_FP[15]) ];
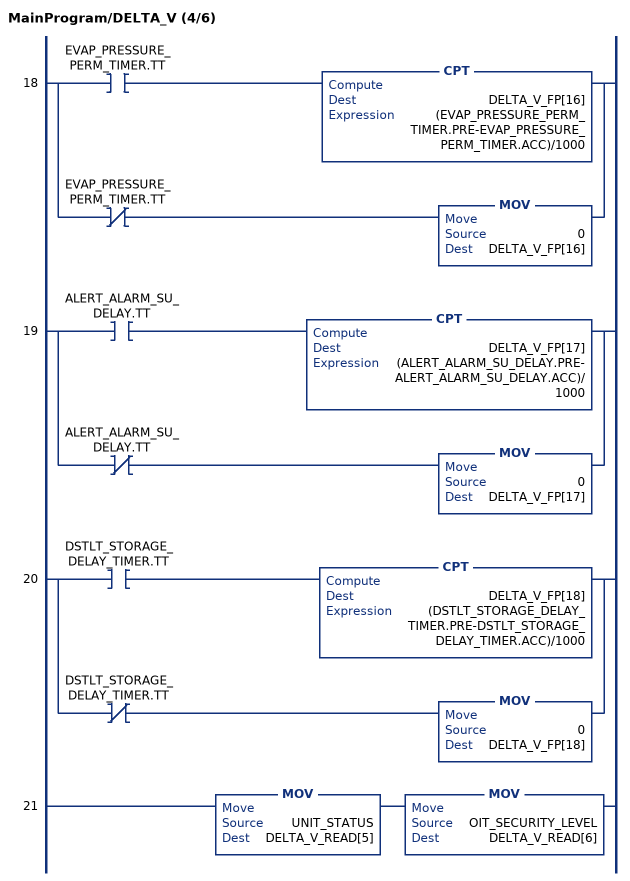
   18: [XIC(EVAP_PRESSURE_PERM_TIMER.TT) CPT(DELTA_V_FP[16],(EVAP_PRESSURE_PERM_TIMER.PRE-EVAP_PRESSURE_PERM_TIMER.ACC)/1000) ,XIO(EVAP_PRESSURE_PERM_TIMER.TT) MOV(0,DELTA_V_FP[16]) ];
   19: [XIC(ALERT_ALARM_SU_DELAY.TT) CPT(DELTA_V_FP[17],(ALERT_ALARM_SU_DELAY.PRE-ALERT_ALARM_SU_DELAY.ACC)/1000) ,XIO(ALERT_ALARM_SU_DELAY.TT) MOV(0,DELTA_V_FP[17]) ];
   20: [XIC(DSTLT_STORAGE_DELAY_TIMER.TT) CPT(DELTA_V_FP[18],(DSTLT_STORAGE_DELAY_TIMER.PRE-DSTLT_STORAGE_DELAY_TIMER.ACC)/1000) ,XIO(DSTLT_STORAGE_DELAY_TIMER.TT) MOV(0,DELTA_V_FP[18]) ];
   21: MOV(UNIT_STATUS,DELTA_V_READ[5])MOV(OIT_SECURITY_LEVEL,DELTA_V_READ[6]);
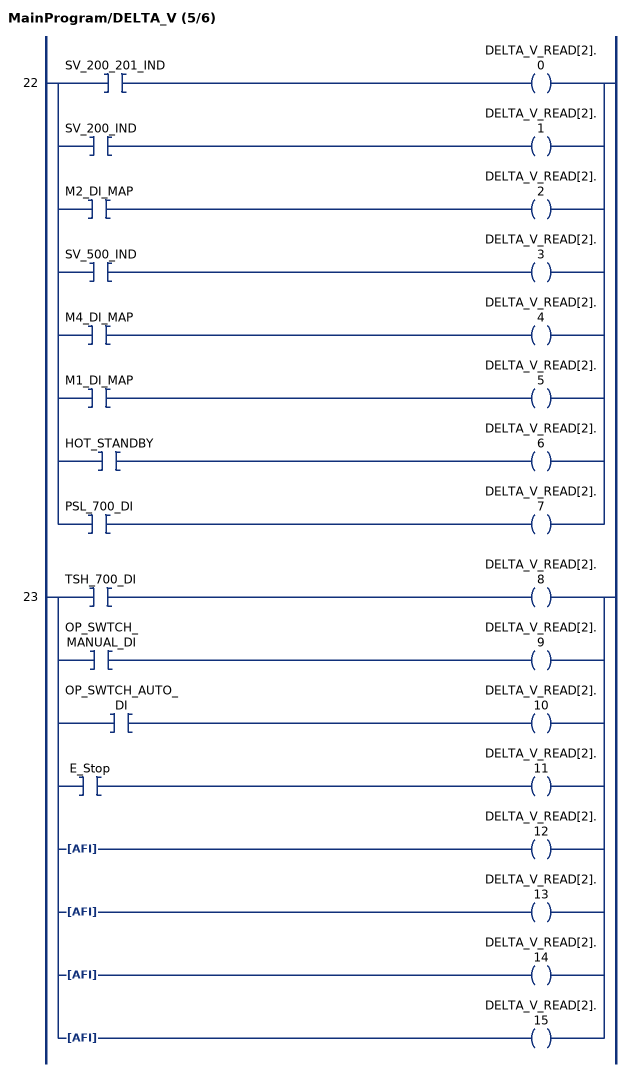
   22: [XIC(SV_200_201_IND) OTE(DELTA_V_READ[2].0) ,XIC(SV_200_IND) OTE(DELTA_V_READ[2].1) ,XIC(M2_DI_MAP) OTE(DELTA_V_READ[2].2) ,XIC(SV_500_IND) OTE(DELTA_V_READ[2].3) ,XIC(M4_DI_MAP) OTE(DELTA_V_READ[2].4) ,XIC(M1_DI_MAP) OTE(DELTA_V_READ[2].5) ,XIC(HOT_STANDBY) OTE(DELTA_V_READ[2].6) ,XIC(PSL_700_DI) OTE(DELTA_V_READ[2].7) ];
   23: [XIC(TSH_700_DI) OTE(DELTA_V_READ[2].8) ,XIC(OP_SWTCH_MANUAL_DI) OTE(DELTA_V_READ[2].9) ,XIC(OP_SWTCH_AUTO_DI) OTE(DELTA_V_READ[2].10) ,XIC(E_Stop) OTE(DELTA_V_READ[2].11) ,AFI() OTE(DELTA_V_READ[2].12) ,AFI() OTE(DELTA_V_READ[2].13) ,AFI() OTE(DELTA_V_READ[2].14) ,AFI() OTE(DELTA_V_READ[2].15) ];
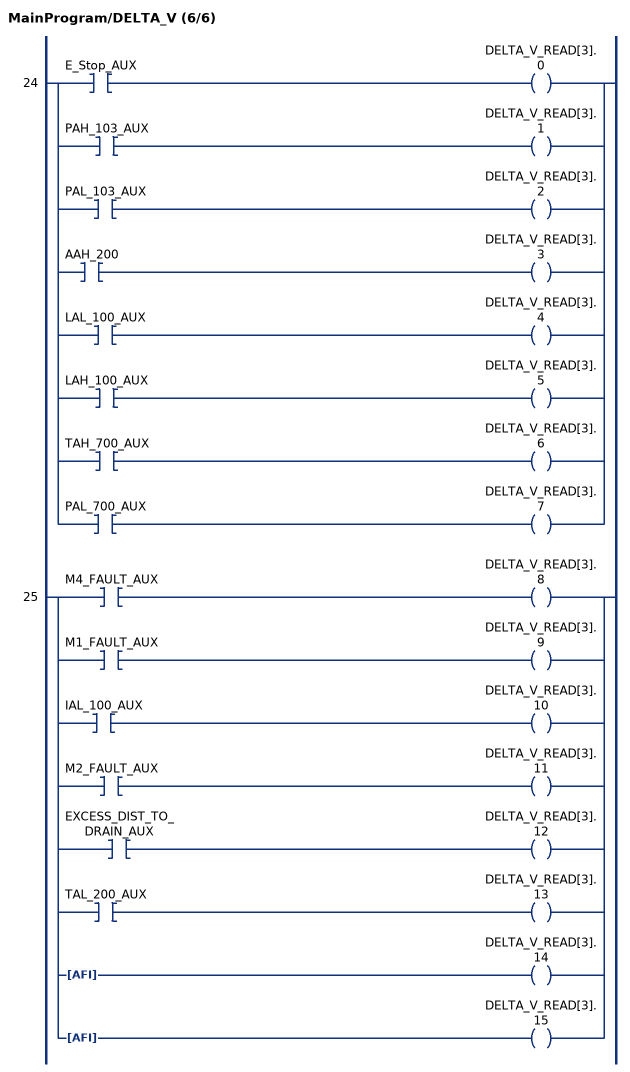
   24: [XIC(E_Stop_AUX) OTE(DELTA_V_READ[3].0) ,XIC(PAH_103_AUX) OTE(DELTA_V_READ[3].1) ,XIC(PAL_103_AUX) OTE(DELTA_V_READ[3].2) ,XIC(AAH_200) OTE(DELTA_V_READ[3].3) ,XIC(LAL_100_AUX) OTE(DELTA_V_READ[3].4) ,XIC(LAH_100_AUX) OTE(DELTA_V_READ[3].5) ,XIC(TAH_700_AUX) OTE(DELTA_V_READ[3].6) ,XIC(PAL_700_AUX) OTE(DELTA_V_READ[3].7) ];
   25: [XIC(M4_FAULT_AUX) OTE(DELTA_V_READ[3].8) ,XIC(M1_FAULT_AUX) OTE(DELTA_V_READ[3].9) ,XIC(IAL_100_AUX) OTE(DELTA_V_READ[3].10) ,XIC(M2_FAULT_AUX) OTE(DELTA_V_READ[3].11) ,XIC(EXCESS_DIST_TO_DRAIN_AUX) OTE(DELTA_V_READ[3].12) ,XIC(TAL_200_AUX) OTE(DELTA_V_READ[3].13) ,AFI() OTE(DELTA_V_READ[3].14) ,AFI() OTE(DELTA_V_READ[3].15) ];
END_ROUTINE

ROUTINE DISTILLATE_LEVEL   (* ladder *)
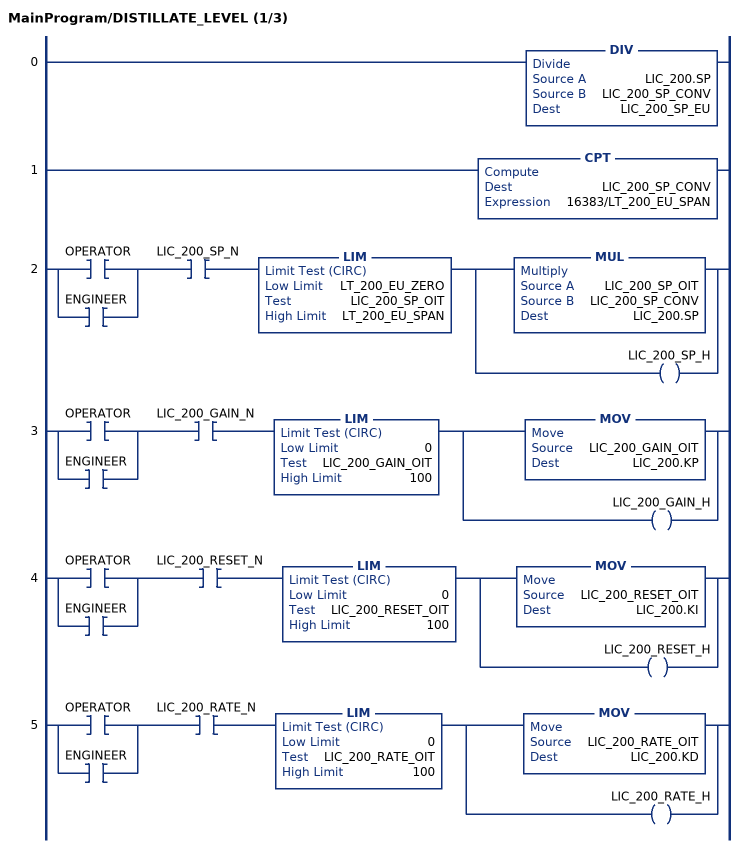
   0: DIV(LIC_200.SP,LIC_200_SP_CONV,LIC_200_SP_EU);
   1: CPT(LIC_200_SP_CONV,16383/LT_200_EU_SPAN);
   2: [XIC(OPERATOR) ,XIC(ENGINEER) ]XIC(LIC_200_SP_N)LIM(LT_200_EU_ZERO,LIC_200_SP_OIT,LT_200_EU_SPAN)[MUL(LIC_200_SP_OIT,LIC_200_SP_CONV,LIC_200.SP) ,OTE(LIC_200_SP_H) ];
   3: [XIC(OPERATOR) ,XIC(ENGINEER) ]XIC(LIC_200_GAIN_N)LIM(0,LIC_200_GAIN_OIT,100)[MOV(LIC_200_GAIN_OIT,LIC_200.KP) ,OTE(LIC_200_GAIN_H) ];
   4: [XIC(OPERATOR) ,XIC(ENGINEER) ]XIC(LIC_200_RESET_N)LIM(0,LIC_200_RESET_OIT,100)[MOV(LIC_200_RESET_OIT,LIC_200.KI) ,OTE(LIC_200_RESET_H) ];
   5: [XIC(OPERATOR) ,XIC(ENGINEER) ]XIC(LIC_200_RATE_N)LIM(0,LIC_200_RATE_OIT,100)[MOV(LIC_200_RATE_OIT,LIC_200.KD) ,OTE(LIC_200_RATE_H) ];
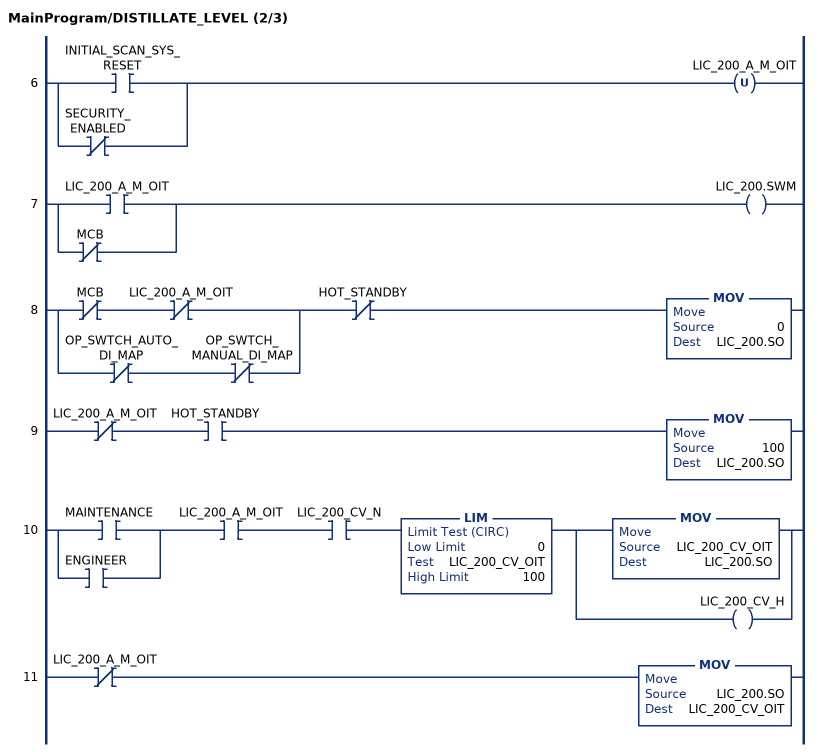
   6: [XIC(INITIAL_SCAN_SYS_RESET) ,XIO(SECURITY_ENABLED) ]OTU(LIC_200_A_M_OIT);
   7: [XIC(LIC_200_A_M_OIT) ,XIO(MCB) ]OTE(LIC_200.SWM);
   8: [XIO(MCB) XIO(LIC_200_A_M_OIT) ,XIO(OP_SWTCH_AUTO_DI_MAP) XIO(OP_SWTCH_MANUAL_DI_MAP) ]XIO(HOT_STANDBY)MOV(0,LIC_200.SO);
   9: XIO(LIC_200_A_M_OIT)XIC(HOT_STANDBY)MOV(100,LIC_200.SO);
   10: [XIC(MAINTENANCE) ,XIC(ENGINEER) ]XIC(LIC_200_A_M_OIT)XIC(LIC_200_CV_N)LIM(0,LIC_200_CV_OIT,100)[MOV(LIC_200_CV_OIT,LIC_200.SO) ,OTE(LIC_200_CV_H) ];
   11: XIO(LIC_200_A_M_OIT)MOV(LIC_200.SO,LIC_200_CV_OIT);
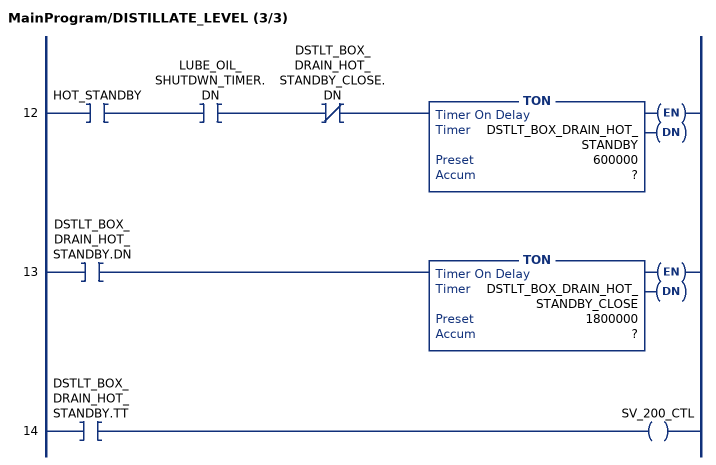
   12: XIC(HOT_STANDBY)XIC(LUBE_OIL_SHUTDWN_TIMER.DN)XIO(DSTLT_BOX_DRAIN_HOT_STANDBY_CLOSE.DN)TON(DSTLT_BOX_DRAIN_HOT_STANDBY,?,?);
   13: XIC(DSTLT_BOX_DRAIN_HOT_STANDBY.DN)TON(DSTLT_BOX_DRAIN_HOT_STANDBY_CLOSE,?,?);
   14: XIC(DSTLT_BOX_DRAIN_HOT_STANDBY.TT)OTE(SV_200_CTL);
END_ROUTINE

ROUTINE DISTILLATE_TEMPERATURE   (* ladder *)
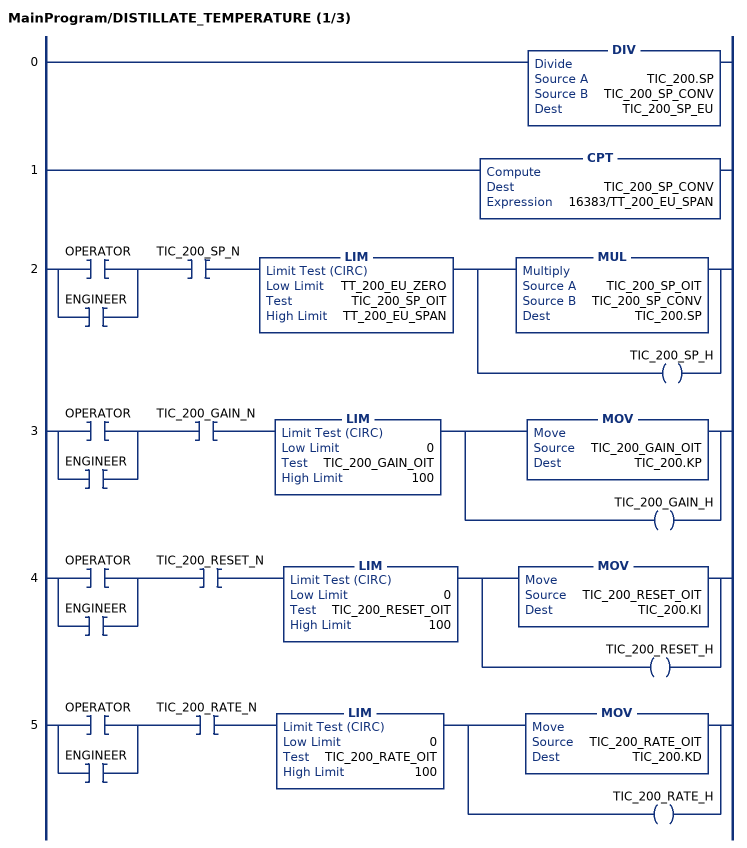
   0: DIV(TIC_200.SP,TIC_200_SP_CONV,TIC_200_SP_EU);
   1: CPT(TIC_200_SP_CONV,16383/TT_200_EU_SPAN);
   2: [XIC(OPERATOR) ,XIC(ENGINEER) ]XIC(TIC_200_SP_N)LIM(TT_200_EU_ZERO,TIC_200_SP_OIT,TT_200_EU_SPAN)[MUL(TIC_200_SP_OIT,TIC_200_SP_CONV,TIC_200.SP) ,OTE(TIC_200_SP_H) ];
   3: [XIC(OPERATOR) ,XIC(ENGINEER) ]XIC(TIC_200_GAIN_N)LIM(0,TIC_200_GAIN_OIT,100)[MOV(TIC_200_GAIN_OIT,TIC_200.KP) ,OTE(TIC_200_GAIN_H) ];
   4: [XIC(OPERATOR) ,XIC(ENGINEER) ]XIC(TIC_200_RESET_N)LIM(0,TIC_200_RESET_OIT,100)[MOV(TIC_200_RESET_OIT,TIC_200.KI) ,OTE(TIC_200_RESET_H) ];
   5: [XIC(OPERATOR) ,XIC(ENGINEER) ]XIC(TIC_200_RATE_N)LIM(0,TIC_200_RATE_OIT,100)[MOV(TIC_200_RATE_OIT,TIC_200.KD) ,OTE(TIC_200_RATE_H) ];
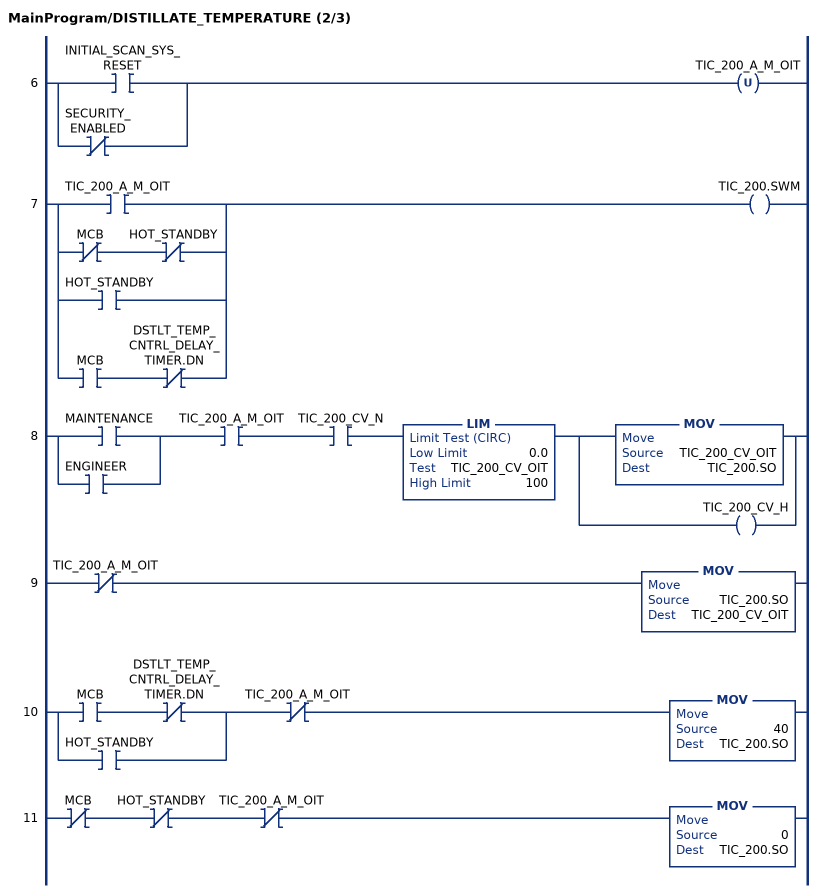
   6: [XIC(INITIAL_SCAN_SYS_RESET) ,XIO(SECURITY_ENABLED) ]OTU(TIC_200_A_M_OIT);
   7: [XIC(TIC_200_A_M_OIT) ,XIO(MCB) XIO(HOT_STANDBY) ,XIC(HOT_STANDBY) ,XIC(MCB) XIO(DSTLT_TEMP_CNTRL_DELAY_TIMER.DN) ]OTE(TIC_200.SWM);
   8: [XIC(MAINTENANCE) ,XIC(ENGINEER) ]XIC(TIC_200_A_M_OIT)XIC(TIC_200_CV_N)LIM(0.0,TIC_200_CV_OIT,100)[MOV(TIC_200_CV_OIT,TIC_200.SO) ,OTE(TIC_200_CV_H) ];
   9: XIO(TIC_200_A_M_OIT)MOV(TIC_200.SO,TIC_200_CV_OIT);
   10: [XIC(MCB) XIO(DSTLT_TEMP_CNTRL_DELAY_TIMER.DN) ,XIC(HOT_STANDBY) ]XIO(TIC_200_A_M_OIT)MOV(40,TIC_200.SO);
   11: XIO(MCB)XIO(HOT_STANDBY)XIO(TIC_200_A_M_OIT)MOV(0,TIC_200.SO);
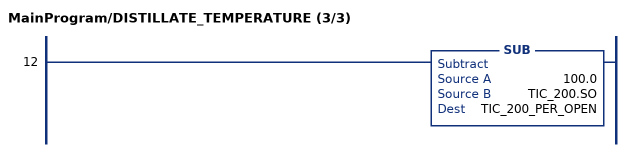
   12: SUB(100.0,TIC_200.SO,TIC_200_PER_OPEN);
END_ROUTINE
